// TIA Portal V21 export
// export: Created 2000-01-01T00:00:00.0000000Z, ExportSetting None
TYPE "UDT_HMI_LowPassFilter"
   STRUCT
      bBypassFilter { ExternalWritable := 'False'} : Bool;   // HMI手动旁路滤波（直通模式）
      bResetCmd { ExternalWritable := 'False'} : Bool;   // HMI手动复位同步触发
      rAlpha { ExternalWritable := 'False'} : Real;   // 滤波系数 Alpha (0.01..1.0，越小越平滑)
      rMaxDeltaPerScan { ExternalWritable := 'False'} : Real;   // 单周期最大允许突变幅值（<=0.0 表示不限制）
      rRawInput { ExternalWritable := 'False'} : Real;   // 状态反馈：原始输入值
      rFilteredOutput { ExternalWritable := 'False'} : Real;   // 状态反馈：滤波后输出值
      bInitialized { ExternalWritable := 'False'} : Bool;   // 状态反馈：已完成冷启动同步
      bError { ExternalWritable := 'False'} : Bool;   // 状态反馈：参数故障标志
      wStatus { ExternalWritable := 'False'} : Word;   // 故障码：16#0000正常, 16#7000未使能, 16#8200系数超范围
   END_STRUCT;
END_TYPE
